Fanuc KAREL source: KT00544.KL

PROGRAM KT00544
%NOLOCKGROUP
VAR
  P1: JOINTPOS
  P2: XYZWPREXT
  OUT: POSITION
BEGIN
    P2.Y = 2.0
  OUT = P1 : P2
END KT00544
